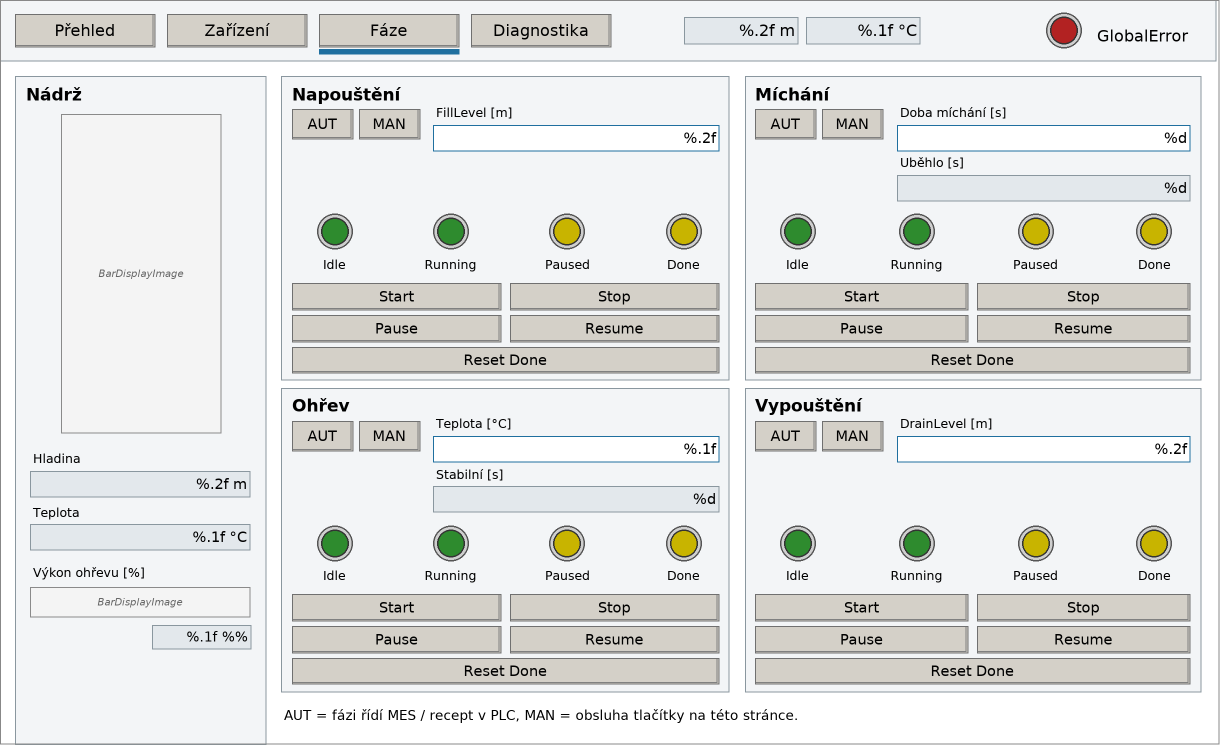
VISUALIZATION Faze  // 1220x745
    Rectangle (0,0 1216x61)
    Button (15,14 140x33), "Přehled"
        OnMouseClick: change screen: Prehled
    Button (167,14 140x33), "Zařízení"
        OnMouseClick: change screen: Zarizeni
    Button (319,14 140x33), "Fáze"
        OnMouseClick: change screen: Faze
    Rectangle (319,49 140x5)
    Button (471,14 140x33), "Diagnostika"
        OnMouseClick: change screen: Diagnostika
    Rectangle (684,17 114x27), "%.2f m", text variable: Global.Tank1.Filling.WaterLevel
    Rectangle (806,17 114x27), "%.1f °C", text variable: Global.Tank1.Heating.WaterTemp
    Lamp1 (1041,10 46x41), variable: Global.Tank1.GlobalError, style: Lamp-Lamp1-Red
    Label (1094,23 126x26), "GlobalError"
    Rectangle (15,76 251x669)
    Label (23,81 65x27), "Nádrž"
    BarDisplayImage (61,114 160x319), value: Global.Tank1.Filling.WaterLevel, style: BarDisplayImage-Gray, scale format: %.1f, scale 0..2
    Label (30,448 66x21), "Hladina"
    Rectangle (30,471 220x26), "%.2f m", text variable: Global.Tank1.Filling.WaterLevel
    Label (30,502 66x21), "Teplota"
    Rectangle (30,524 220x26), "%.1f °C", text variable: Global.Tank1.Heating.WaterTemp
    Label (30,562 142x21), "Výkon ohřevu [%]"
    BarDisplayImage (30,587 220x30), value: Global.Tank1.Heater.State.HeatingOut, style: BarDisplayImage-Gray, scale format: %.1f, scale 0..100
    Rectangle (152,625 99x24), "%.1f %%", text variable: Global.Tank1.Heater.State.HeatingOut
    Rectangle (281,76 448x304)
    Label (289,81 122x27), "Napouštění"
    Button (292,109 61x30), "AUT", colour toggle: Global.Tank1.Filling.State.AutCtrl
        tap Global.Tank1.Filling.Cmd.AutCtrl
    Button (359,109 61x30), "MAN", colour toggle: Global.Tank1.Filling.State.ManCtrl
        tap Global.Tank1.Filling.Cmd.ManCtrl
    Label (433,102 117x21), "FillLevel [m]"
    Rectangle (433,125 286x26), "%.2f", text variable: Global.Tank1.Filling.ParamFillLevel
        OnMouseClick: write the text variable via Default
    Lamp1 (312,211 46x41), variable: Global.Tank1.Filling.State.Idle, style: Lamp-Lamp1-Green
    Label (289,254 91x21), "Idle"
    Lamp1 (428,211 46x41), variable: Global.Tank1.Filling.State.Running, style: Lamp-Lamp1-Green
    Label (405,254 91x21), "Running"
    Lamp1 (544,211 46x41), variable: Global.Tank1.Filling.State.Paused, style: Lamp-Lamp1-Yellow
    Label (522,254 91x21), "Paused"
    Lamp1 (661,211 46x41), variable: Global.Tank1.Filling.State.Done, style: Lamp-Lamp1-Yellow
    Label (638,254 91x21), "Done"
    Button (292,283 209x27), "Start", colour toggle: Global.Tank1.Filling.State.Running
        tap Global.Tank1.Filling.Cmd.StartMan
    Button (510,283 209x27), "Stop"
        tap Global.Tank1.Filling.Cmd.StopMan
    Button (292,315 209x27), "Pause", colour toggle: Global.Tank1.Filling.State.Paused
        tap Global.Tank1.Filling.Cmd.PauseMan
    Button (510,315 209x27), "Resume"
        tap Global.Tank1.Filling.Cmd.ResumeMan
    Button (292,347 427x26), "Reset Done", colour toggle: Global.Tank1.Filling.State.Done
        tap Global.Tank1.Filling.Cmd.ResetDone
    Rectangle (745,76 456x304)
    Label (752,81 87x27), "Míchání"
    Button (755,109 61x30), "AUT", colour toggle: Global.Tank1.Mixing.State.AutCtrl
        tap Global.Tank1.Mixing.Cmd.AutCtrl
    Button (822,109 61x30), "MAN", colour toggle: Global.Tank1.Mixing.State.ManCtrl
        tap Global.Tank1.Mixing.Cmd.ManCtrl
    Label (897,102 142x21), "Doba míchání [s]"
    Rectangle (897,125 293x26), "%d", text variable: Global.Tank1.Mixing.ParamTimeSec
        OnMouseClick: write the text variable via Default
    Label (897,152 92x21), "Uběhlo [s]"
    Rectangle (897,175 293x26), "%d", text variable: Global.Tank1.Mixing.ElapsedTimeSec
    Lamp1 (775,211 46x41), variable: Global.Tank1.Mixing.State.Idle, style: Lamp-Lamp1-Green
    Label (752,254 91x21), "Idle"
    Lamp1 (894,211 46x41), variable: Global.Tank1.Mixing.State.Running, style: Lamp-Lamp1-Green
    Label (871,254 91x21), "Running"
    Lamp1 (1013,211 46x41), variable: Global.Tank1.Mixing.State.Paused, style: Lamp-Lamp1-Yellow
    Label (990,254 91x21), "Paused"
    Lamp1 (1131,211 46x41), variable: Global.Tank1.Mixing.State.Done, style: Lamp-Lamp1-Yellow
    Label (1109,254 91x21), "Done"
    Button (755,283 213x27), "Start", colour toggle: Global.Tank1.Mixing.State.Running
        tap Global.Tank1.Mixing.Cmd.StartMan
    Button (977,283 213x27), "Stop"
        tap Global.Tank1.Mixing.Cmd.StopMan
    Button (755,315 213x27), "Pause", colour toggle: Global.Tank1.Mixing.State.Paused
        tap Global.Tank1.Mixing.Cmd.PauseMan
    Button (977,315 213x27), "Resume"
        tap Global.Tank1.Mixing.Cmd.ResumeMan
    Button (755,347 435x26), "Reset Done", colour toggle: Global.Tank1.Mixing.State.Done
        tap Global.Tank1.Mixing.Cmd.ResetDone
    Rectangle (281,388 448x304)
    Label (289,392 65x27), "Ohřev"
    Button (292,421 61x30), "AUT", colour toggle: Global.Tank1.Heating.State.AutCtrl
        tap Global.Tank1.Heating.Cmd.AutCtrl
    Button (359,421 61x30), "MAN", colour toggle: Global.Tank1.Heating.State.ManCtrl
        tap Global.Tank1.Heating.Cmd.ManCtrl
    Label (433,413 109x21), "Teplota [°C]"
    Rectangle (433,436 286x26), "%.1f", text variable: Global.Tank1.Heating.ParamReqTemp
        OnMouseClick: write the text variable via Default
    Label (433,464 109x21), "Stabilní [s]"
    Rectangle (433,486 286x26), "%d", text variable: Global.Tank1.Heating.fTime
    Lamp1 (312,523 46x41), variable: Global.Tank1.Heating.State.Idle, style: Lamp-Lamp1-Green
    Label (289,565 91x21), "Idle"
    Lamp1 (428,523 46x41), variable: Global.Tank1.Heating.State.Running, style: Lamp-Lamp1-Green
    Label (405,565 91x21), "Running"
    Lamp1 (544,523 46x41), variable: Global.Tank1.Heating.State.Paused, style: Lamp-Lamp1-Yellow
    Label (522,565 91x21), "Paused"
    Lamp1 (661,523 46x41), variable: Global.Tank1.Heating.State.Done, style: Lamp-Lamp1-Yellow
    Label (638,565 91x21), "Done"
    Button (292,594 209x27), "Start", colour toggle: Global.Tank1.Heating.State.Running
        tap Global.Tank1.Heating.Cmd.StartMan
    Button (510,594 209x27), "Stop"
        tap Global.Tank1.Heating.Cmd.StopMan
    Button (292,626 209x27), "Pause", colour toggle: Global.Tank1.Heating.State.Paused
        tap Global.Tank1.Heating.Cmd.PauseMan
    Button (510,626 209x27), "Resume"
        tap Global.Tank1.Heating.Cmd.ResumeMan
    Button (292,658 427x26), "Reset Done", colour toggle: Global.Tank1.Heating.State.Done
        tap Global.Tank1.Heating.Cmd.ResetDone
    Rectangle (745,388 456x304)
    Label (752,392 122x27), "Vypouštění"
    Button (755,421 61x30), "AUT", colour toggle: Global.Tank1.Draining.State.AutCtrl
        tap Global.Tank1.Draining.Cmd.AutCtrl
    Button (822,421 61x30), "MAN", colour toggle: Global.Tank1.Draining.State.ManCtrl
        tap Global.Tank1.Draining.Cmd.ManCtrl
    Label (897,413 125x21), "DrainLevel [m]"
    Rectangle (897,436 293x26), "%.2f", text variable: Global.Tank1.Draining.ParamDrainLevel
        OnMouseClick: write the text variable via Default
    Lamp1 (775,523 46x41), variable: Global.Tank1.Draining.State.Idle, style: Lamp-Lamp1-Green
    Label (752,565 91x21), "Idle"
    Lamp1 (894,523 46x41), variable: Global.Tank1.Draining.State.Running, style: Lamp-Lamp1-Green
    Label (871,565 91x21), "Running"
    Lamp1 (1013,523 46x41), variable: Global.Tank1.Draining.State.Paused, style: Lamp-Lamp1-Yellow
    Label (990,565 91x21), "Paused"
    Lamp1 (1131,523 46x41), variable: Global.Tank1.Draining.State.Done, style: Lamp-Lamp1-Yellow
    Label (1109,565 91x21), "Done"
    Button (755,594 213x27), "Start", colour toggle: Global.Tank1.Draining.State.Running
        tap Global.Tank1.Draining.Cmd.StartMan
    Button (977,594 213x27), "Stop"
        tap Global.Tank1.Draining.Cmd.StopMan
    Button (755,626 213x27), "Pause", colour toggle: Global.Tank1.Draining.State.Paused
        tap Global.Tank1.Draining.Cmd.PauseMan
    Button (977,626 213x27), "Resume"
        tap Global.Tank1.Draining.Cmd.ResumeMan
    Button (755,658 435x26), "Reset Done", colour toggle: Global.Tank1.Draining.State.Done
        tap Global.Tank1.Draining.Cmd.ResetDone
    Label (281,704 682x23), "AUT = fázi řídí MES / recept v PLC, MAN = obsluha tlačítky na této stránce."
END_VISUALIZATION

(* stored: Version 1.1.0.1, ProductVersion 3.1.4026.21
   Visu Faze: Id {66f97671-98e5-42d9-9654-6f663eac1bc2} *)
